(*
SPDX-FileCopyrightText: © 2026 Oleksandr Tiutyk <trofimich@gmail.com>
SPDX-License-Identifier: MIT
License: https://opensource.org/license/mit
*)

(*
Checks that FB_reinit preserves scaling limits and fallback references in range converters.

Exercises FB_reinit in place on StaticRangeAnalogValueConverter and DynamicRangeAnalogValueConverter;
copy-code relocation requires a TwinCAT runtime online-change check.
*)

{attribute 'no_assign'}
{attribute 'no_explicit_call' := 'do not call this function block directly'}
FUNCTION_BLOCK ConverterOnlineChangeLifecycleTest EXTENDS TOF_Testing.SingleCycleTest
VAR_STAT
	{attribute 'hide'}
	_ClassName : STRING := __POUNAME();
END_VAR

(* Verifies static limits, live dynamic references, and zero fallback references across FB_reinit. *)
METHOD PROTECTED ExecuteTest
VAR
	minAnalog : LREAL := 0.0;
	maxAnalog : LREAL := 100.0;
	minRaw : TOF_Devices_IO.RAW_ANALOG_VALUE := TOF_Devices_IO.RawAnalogValues.FromInt16(value := 0);
	maxRaw : TOF_Devices_IO.RAW_ANALOG_VALUE := TOF_Devices_IO.RawAnalogValues.FromInt16(value := 1000);
	invalidMaxRaw : REFERENCE TO TOF_Devices_IO.RAW_ANALOG_VALUE;
	staticConverter : TOF_Devices_IO.StaticRangeAnalogValueConverter(
		minAnalogValue := 0.0,
		maxAnalogValue := 100.0,
		minRawValue := minRaw,
		maxRawValue := maxRaw
	);
	dynamicConverter : TOF_Devices_IO.DynamicRangeAnalogValueConverter(
		minAnalogValue := minAnalog,
		maxAnalogValue := maxAnalog,
		minRawValue := minRaw,
		maxRawValue := maxRaw
	);
	fallbackConverter : TOF_Devices_IO.DynamicRangeAnalogValueConverter(
		minAnalogValue := minAnalog,
		maxAnalogValue := maxAnalog,
		minRawValue := minRaw,
		maxRawValue := invalidMaxRaw
	);
	rawResult : TOF_Devices_IO.RAW_ANALOG_VALUE;
	reinitialized : BOOL;
END_VAR
reinitialized := staticConverter.FB_reinit()
	AND_THEN dynamicConverter.FB_reinit()
	AND_THEN fallbackConverter.FB_reinit();
Assert.ThatBool(
	actual := reinitialized,
	message := "Converter FB_reinit calls must return TRUE"
).IsTrue();

Assert.ThatLongReal(
	actual := staticConverter.MaxAnalogValue,
	message := "Static converter must retain configured analog maximum after FB_reinit"
).ToBe(expected := 100.0, tolerance := 0.001);

rawResult := staticConverter.ConvertAnalogValueToRawValue(
	analogValue := 50.0,
	rawValueType := TOF_Devices_IO.RAW_ANALOG_VALUE_TYPE.INT16
);
Assert.ThatInt(
	actual := rawResult.Int16,
	message := "Static converter must scale accurately after FB_reinit"
).ToBe(expected := 500);

rawResult := staticConverter.ConvertAnalogValueToRawValue(
	analogValue := 150.0,
	rawValueType := TOF_Devices_IO.RAW_ANALOG_VALUE_TYPE.INT16
);
Assert.ThatInt(
	actual := rawResult.Int16,
	message := "Static converter must keep upper raw clamping after FB_reinit"
).ToBe(expected := 1000);

maxAnalog := 200.0;
rawResult := dynamicConverter.ConvertAnalogValueToRawValue(
	analogValue := 50.0,
	rawValueType := TOF_Devices_IO.RAW_ANALOG_VALUE_TYPE.INT16
);
Assert.ThatInt(
	actual := rawResult.Int16,
	message := "Dynamic converter must continue tracking referenced limits after FB_reinit"
).ToBe(expected := 250);

rawResult := fallbackConverter.ConvertAnalogValueToRawValue(
	analogValue := 50.0,
	rawValueType := TOF_Devices_IO.RAW_ANALOG_VALUE_TYPE.INT16
);
Assert.ThatInt(
	actual := rawResult.Int16,
	message := "Dynamic converter must preserve zero fallback limits after FB_reinit"
).ToBe(expected := 0);
END_METHOD

// Borrows the concrete class name. Callers must not modify it.
{attribute 'monitoring' := 'call'}
PROPERTY ClassName : REFERENCE TO STRING
GET
ClassName REF= _ClassName;
END_GET
END_PROPERTY

// Borrows the compiler-initialized namespace name. Callers must not modify it.
{attribute 'monitoring' := 'call'}
PROPERTY NamespaceName : REFERENCE TO STRING
GET
NamespaceName REF= CurrentNamespace.Name;
END_GET
END_PROPERTY

// Reports the concrete instance size in bytes.
{attribute 'monitoring' := 'call'}
PROPERTY SelfSize : ULINT
GET
SelfSize := XSIZEOF(THIS^);
END_GET
END_PROPERTY

END_FUNCTION_BLOCK

(* stored: Version 1.1.0.1
   POU ConverterOnlineChangeLifecycleTest: Id {5d2554b8-6d83-4347-8980-d85ec37133ec}, SpecialFunc None
   Method ExecuteTest: Id {879f1745-04fd-45e1-9e71-c564ebcc5281}
   Property ClassName: Id {c8e7f6b1-40de-4fee-9bea-8b612decafc9}
   Get Get: Id {88129ece-9a7c-4479-9698-e16332ed4b63}
   Property NamespaceName: Id {ccb1e945-d8cb-4b8e-b31e-ca8d82ec8d92}
   Get Get: Id {8234a1fc-9e2c-488b-b8c7-b2bf429b39a3}
   Property SelfSize: Id {c9e04095-6d74-4849-8af4-5b9b6f11ac4e}
   Get Get: Id {7284b187-2c6e-4f02-9313-715c484d2052} *)
